(*
SPDX-FileCopyrightText: © 2026 Oleksandr Tiutyk <trofimich@gmail.com>
SPDX-License-Identifier: MIT
License: https://opensource.org/license/mit
*)

(*
Internal target used by Workflow.FB_reinit to update direct workflow associations after relocation.

Implementations update _Workflow only when a direct association was already set so inherited parent-resolved
associations remain untouched.
*)
{attribute 'hide'}
INTERFACE INTERNAL IWorkflowAssociationTarget EXTENDS TOF_Core.IObject

(* Updates a direct workflow association after the owning workflow relocated during online change. *)
METHOD RebindWorkflow
VAR_INPUT
	workflow : IWorkflow;
END_VAR
END_METHOD

END_INTERFACE

(* stored: Version 1.1.0.1
   Itf IWorkflowAssociationTarget: Id {0325a656-32cd-4f55-9d85-2d799046441f}
   Method RebindWorkflow: Id {36bb76f6-18c6-4119-922e-6887e572af7e} *)
